(* IEC 61131-3 sources: llm-plc-st-eval/data/definitivo/gemini-3.1-pro-preview/B8/zero_shot, 3 files *)

(* ---- ejec_1.st ---- *)
```iecst
FUNCTION_BLOCK FB_Puerta
VAR_INPUT
    puertaAbierta : BOOL; (* Señal de estado de la puerta (TRUE = abierta) *)
    reset : BOOL;         (* Señal para reiniciar el contador y apagar el aviso *)
END_VAR

VAR_OUTPUT
    aviso : BOOL;         (* Indicador de alarma por 5 o más aperturas *)
    nAperturas : INT;     (* Registro del número de aperturas acumuladas *)
END_VAR

VAR
    flancoApertura : R_TRIG; (* Instancia para detectar el flanco de subida *)
END_VAR

(* Detección de la transición de FALSE a TRUE en la señal de la puerta *)
flancoApertura(CLK := puertaAbierta);

(* Lógica de reinicio y conteo de aperturas *)
IF reset THEN
    nAperturas := 0;
ELSIF flancoApertura.Q THEN
    nAperturas := nAperturas + 1;
END_IF;

(* Activación del aviso si se alcanzan 5 o más aperturas *)
aviso := (nAperturas >= 5);

END_FUNCTION_BLOCK
```

(* ---- ejec_2.st ---- *)
```iecst
FUNCTION_BLOCK FB_Puerta
VAR_INPUT
    puertaAbierta : BOOL; (* Señal de estado de la puerta de seguridad *)
    reset : BOOL;         (* Pone a cero el contador y apaga el aviso *)
END_VAR

VAR_OUTPUT
    aviso : BOOL;         (* TRUE si se acumulan 5 o más aperturas *)
    nAperturas : INT;     (* Número acumulado de aperturas *)
END_VAR

VAR
    flancoApertura : R_TRIG; (* Detector de flanco de subida estándar IEC *)
END_VAR

(* Detectar transición de FALSE a TRUE en la señal de la puerta *)
flancoApertura(CLK := puertaAbierta);

(* Lógica de reinicio o incremento del contador *)
IF reset THEN
    nAperturas := 0;
ELSIF flancoApertura.Q THEN
    nAperturas := nAperturas + 1;
END_IF;

(* Evaluación de la salida de aviso (se desactiva automáticamente al resetear nAperturas) *)
aviso := (nAperturas >= 5);

END_FUNCTION_BLOCK
```

(* ---- ejec_3.st ---- *)
```iecst
FUNCTION_BLOCK FB_Puerta
VAR_INPUT
    puertaAbierta : BOOL; // Señal de estado de la puerta (TRUE = abierta)
    reset : BOOL;         // Señal para reiniciar el contador y apagar el aviso
END_VAR

VAR_OUTPUT
    aviso : BOOL;         // Indicador de 5 o más aperturas
    nAperturas : INT;     // Registro del número de aperturas
END_VAR

VAR
    flancoApertura : R_TRIG; // Instancia para detectar el flanco de subida
END_VAR

// Detección de la transición de FALSE a TRUE en la entrada puertaAbierta
flancoApertura(CLK := puertaAbierta);

// Lógica de reinicio y conteo de aperturas
IF reset THEN
    nAperturas := 0;
ELSIF flancoApertura.Q THEN
    nAperturas := nAperturas + 1;
END_IF;

// Evaluación de la salida de aviso (se desactiva automáticamente al resetear)
aviso := (nAperturas >= 5);

END_FUNCTION_BLOCK
```
